DATA_BLOCK "S12Probe"
{ S7_Optimized_Access := 'TRUE' }
VERSION : 0.1
NON_RETAIN
   VAR
      Stage : DInt;
      Ready : Bool;
      Initialized : Bool;
      Scans : UDInt;
      MonoSec : LReal;
      MaxDeltaSec : LReal;
      BadDelta : UDInt;
      RuntimeMem : LReal;
      ClockStart : DTL;
      ClockNow : DTL;
      ClockRc : Int;
      BoolTrue : Bool;
      BoolFalse : Bool;
      IntMin : Int;
      IntMax : Int;
      DIntMin : DInt;
      DIntMax : DInt;
      UIntMax : UInt;
      UDIntMax : UDInt;
      RealValue : Real;
      LRealValue : LReal;
      TimeValue : Time;
      NegativeTime : Time;
      LongMin : LInt;
      LongMax : LInt;
      UnsignedMax : ULInt;
      BeyondJsonExact : ULInt;
      StampDtl : DTL;
      StampLdt : LDT;
      StampDt : Date_And_Time;
      Text254 : String[254];
      Text255 : WString[255];
      Text480 : WString[480];
      Text254Length : DInt;
      Text255Length : DInt;
      Text480Length : DInt;
      WideConcat : WString[480];
      WideTail : WString[3];
      EscapedText : String[32];
      UnicodeText : WString[32];
      LowerArray : Array[-2..2] of DInt;
      EnumWitness : DInt;
      WriteWitness : DInt;
   END_VAR
BEGIN
END_DATA_BLOCK
